(* IEC 61131-3 sources: Elmo_Master/Lasal_PRG/Welcon8Axis_EtherCAT_Test_With_RobotAxis/Network/HW_Network, 1 file *)

(* ---- ONE_HW_Network_Table.st ---- *)
#define OBJECTS_CONFIG

//Define part of class _SyncMeasure
#define _SYNCM_PLLLOCK_MASK 2#11110000
#define _SYNCM_PLLLOCK      2#10100000

#define _SYNCM_PLLLOCK_MASK_MASTER 2#11000000
#define _SYNCM_PLLLOCK_MASTER      2#10000000

#define _SYNCM_PLLLOCK_MASK_OWN 2#00110000
#define _SYNCM_PLLLOCK_OWN      2#00100000

#define _SYNCM_PLL_DELTAREG_ENABLE   2#01001000
#define _SYNCM_PLL_DELTAREG_DISABLE  2#01000000

#define _SYNCM_25US 2500 // [10 ns]
#define _SYNCM_50US 5000 // [10 ns]

// #define _SYNCM_DEBUG
#include "..\..\source\interfaces\lsl_st_pll.h"
#include "..\..\Source\BusInterface.h"
//Define part of class _SyncMeasureECAT
#define _SYNCMCAT_MAX_FILTER_SIZE 100

//#define _SYNCMECAT_DEBUG

#define _SYNCMECAT_FilterSize_LL_Measure_Delta   150
#define _SYNCMECAT_FilterSize_LLFP_Offset         25
#define _SYNCMECAT_FilterSize_LL_Roundtrip       500
#define _SYNCMECAT_FilterSize_RCLL_Offset         10
#define _SYNCMECAT_FilterSize_Deltatime           10
#define _SYNCMECAT_FilterSize_Gradient            30
#define _SYNCMECAT_FilterSize_Corr_Steig          80

#define _SYNCMECAT_DCSlvM_AdjustLevel             1//10 //ns

#define _SYNCMECAT_SyncStart_CorrFactorUp        100
#define _SYNCMECAT_SyncStart_CorrFactorDown       50

#define _SYNCMECAT_SyncStart_CorrFactorUp_fine     1
#define _SYNCMECAT_SyncStart_CorrFactorDown_fine   1

#define _SYNCMECAT_SyncStart_DistFactUp        25000
#define _SYNCMECAT_SyncStart_DistFactDown      25000
#include "..\..\Class\ECAT_Master_Base\ECAT_Master_Base.h"
#include "..\..\Class\_SyncMeasureECAT\_64BitTimestamp.h"
//Define part of class BusInterfaceSDIASInternal
#define BUSIF_INTERNAL_MAX_NR_DO 100

// Defines for Mutex Generation
#define INTERNAL_STR_MUTEX_NAME_SEPERATOR ".."
#define INTERNAL_MUTEX_NAME_END_LENGTH 5
#define INTERNAL_MUTEX_NAME_MAX_LENGTH 32
#include "..\..\Source\interfaces\lsl_st_mt.h"
#include "..\..\Class\HwControl\HwControl.h"
#include "..\..\Source\interfaces\lsl_st_hardwaretree.h"
//Define part of class ECAT_Slave_Base
#define ECAT_SB_SDO_LOCK                    16#A1B2C3D4
#define ECAT_SB_SDO_FREE                    16#E5F60718

#define ECAT_SB_VENDORID_SIGMATEK           16#000088FA

//CoE Communication area
#define ECAT_SB_INDEX_DEVICE_TYPE           16#1000 //mandatory
#define ECAT_SB_SUBINDEX_DEVICE_TYPE              0

#define ECAT_SB_INDEX_DEVICE_NAME           16#1008 //optional
#define ECAT_SB_SUBINDEX_DEVICE_NAME              0

#define ECAT_SB_INDEX_HARDWARE_VERSION      16#1009 //optional
#define ECAT_SB_SUBINDEX_HARDWARE_VERSION         0

#define ECAT_SB_INDEX_SOFTWARE_VERSION      16#100A //optional
#define ECAT_SB_SUBINDEX_SOFTWARE_VERSION         0

#define ECAT_SB_INDEX_IDENTITY_OBJECT       16#1018 //mandatory
#define ECAT_SB_SUBINDEX_IDENTITY_OBJECT          0

#define ECAT_SB_DEFAULT_SDO_TIMEOUT         2000

#define ECAT_SB_PHYSICAL_START_ADRESS        1001
#include "..\..\Class\ECAT_Slave_Base\ECAT_Slave_Base.h"
#include "..\..\Source\interfaces\lsl_st_ecatm.h"
//Define part of class ECAT_DS402Base
// As defined in ETG.6010 D (R) V1.1.0

// PDO idx
#define ECAT_DS402BASE_IDX_CONTROLWORD  0x6040
#define ECAT_DS402BASE_IDX_STATUSWORD   0x6041

#define ECAT_DS402BASE_IDX_SETSPEED     0x60FF
#define ECAT_DS402BASE_IDX_ACTSPEED     0x606C

#define ECAT_DS402BASE_IDX_SETPOS       0x607A
#define ECAT_DS402BASE_IDX_ACTPOS       0x6064

#define ECAT_DS402BASE_IDX_ACTTORQUE    0x6077
#define ECAT_DS402BASE_IDX_SETTORQUE    0x6071

#define ECAT_DS402BASE_IDX_ACTXW        0x60F4
#include "..\..\Source\DriveSafetyIF.h"
//Define part of class ECAT_Master_Base
#define ECATM_MAX_NO_TASKS 5
#define ECATM_INC_CYC_CALLBACKS 5

#define ECATM_STR_ENI_FILE    "C:/lslsys/hwoutput.conf"      //Standard path of ENI-File

#define ECATM_MAX_VALUE_MISSING_FRAME_BEHAVIOUR 31
#define ECATM_MAX_SIZE_FRAME_ERROR_LOGBUFFER    50

#define ECATM_THREAD_PRIO_DISABLE               10 // Background
#define ECATM_THREAD_STACKSIZE              0x4000
#include "..\..\Source\interfaces\lsl_st_systrace.h"
#include "..\..\Source\interfaces\lsl_st_gpio.h"
#include "..\..\Source\interfaces\lsl_st_mediaplayer.h"
#include "..\..\Source\interfaces\lsl_st_pci.h"
#include "..\..\Source\interfaces\lsl_st_powermanagement.h"
#include "..\..\Source\interfaces\lsl_st_pwm.h"
#include "..\..\source\interfaces\lsl_st_spi.h"
#include "..\..\Source\interfaces\lsl_st_sysinfo.h"
#include "..\..\Source\interfaces\lsl_st_x_ram.h"
#include "..\..\Class\HwControl\watchdog.h"
#include "..\..\Class\HwControl\_HWKScope.h"
#include "..\..\Class\HwControl\HwControlParameters.h"
#include <.\lsl_st_mt.h>
//Define part of class SafetyUDP
#define SAFETY_UDP_MAX_SOCKETS                6     // Max number of socket

#define SAFETY_UDP_CLT_SEND_OK                0    // Send ok
#define SAFETY_UDP_CLT_INVALID_HANDLE        -1    // Invalid handle
#define SAFETY_UDP_CLT_NOT_OPEN              -2    // Socket is not open
#define SAFETY_UDP_CLT_SEND_FAILED           -3    // Send failed
#define SAFETY_UDP_CLT_SEND_BUFFER_FULL      -4    // Send buffer is full
#define SAFETY_UDP_CLT_DATA_TO_BIG           -5    // Data to big

#define SAFETY_UDP_MAXIMUM_SEGMENT_SIZE    1452    // Maximum of user data

#define SAFETY_UDP_TIMEOUT_OPENSOCKET    (1000)    //timeout for opening socket

#define SAFETY_UDP_RECEIVE_TIMEOUT          800

#define SAFETY_UDP_TX_BUFFER_SIZE          1024
//Define part of class SafetyManager
#define SM_LogBufferSize 1000
#define SM_MaxObjNameLen  256
#include "..\..\Class\SafetyManager\SafetyManager.h"
#include "..\..\Source\interfaces\lsl_st_safetydll.h"
//Define part of class SafetyRoutingTables
#define SRT_MAXIDX 15 // Currently there are 2 Tables for each Eni File / EtherMaster
//Define part of class SdiasManager
#define SDIAS_SDO_MAX_LENGTH              128
#define SDIAS_SDO_RINGBUFFER_NO            64
#define SDIAS_SDO_CHANNEL_NO                3   // fixed in the VI hardware to be 3

// watchdog trigger interval (after 130ms of no trigger the SDIAS HW goes into reset again and takes at least another 10ms to be ready again)
#define SDIAS_WATCHDOG_TRIGGER_TIME        40

// time needed by sdias modules to start up after the watchdog is triggered the first time in ms
#define SDIAS_HARDWARE_STARTUP_TIME        15

// sdias manager needs 2 ticks to handle event for read task (measure sync time)
#define SDIAS_SYNC_MEASURE_TICKS            2

// after activating the PLL SyncOut it takes 3 cycles until the SDIAS sync can be injected
#define SDIAS_CYCLES_WAIT_AFTER_SYNC_ENABLE 3

// wait 1 bus cycle at start to get valid numbers in the task info
#define SDIAS_TASKINFO_READY_TICKS          1

// time to wait (in ms) until other tasks in the same or lower priority than post init have done their stuff
#define SDIAS_WAIT_TIME_IN_POST_INIT        1

#define SIZE_PER_SDIAS_CLIENT               16#0400

// for far memory accesses: 1 module can hold maximum 256 1K blocks (0-255)
#define SDIAS_1K_BLOCK_NO                       256

// far memory accesses maximum length in bytes
#define SDIAS_MAX_SIZE_FAR_MEM_ACCESS           127

#define SDIAS_OFFSET_HW_CONFIG              16#FF00
#define SDIAS_OFFSET_TASK_EVENT_IDS         16#FF10
#define SDIAS_OFFSET_FEATURE_INFO           16#FF18
#define SDIAS_OFFSET_APPLI_LED_STATES       16#FF20
#define SDIAS_OFFSET_SYNC_INJECTION_CFG     16#FF3D
#define SDIAS_OFFSET_TRIGGER_UNIT_SETUP_0   16#FF41
#define SDIAS_OFFSET_TRIGGER_UNIT_SETUP_1   16#FF45
#define SDIAS_OFFSET_TASK_START_CFG_0       16#FF60
#define SDIAS_OFFSET_TASK_CONFIG_0          16#FF86
#define SDIAS_OFFSET_TASK_CONFIG_1          16#FF96
#define SDIAS_OFFSET_TASK_INFO_1            16#FF94
#define SDIAS_OFFSET_TASK_HANDSHAKE_1       16#FF9B
#define SDIAS_OFFSET_TASK_DURATION_TIME_1   16#FF9C
#define SDIAS_OFFSET_TASK_DURATION_TIME_2   16#FFAC
#define SDIAS_OFFSET_TASK_CONFIG_2          16#FFA6

#define SDIAS_RETRIES_ALLOWED         2

// mask to get global error flag out of message counter byte of SDO responses
#define SDIAS_MASK_GLOBAL_ERROR_FLAG        16#80

// mask to get message counter out of message counter byte of SDO responses
#define SDIAS_MASK_MESSAGE_COUNTER          16#3F

#define SDIAS_EVENT_MASK_ID_SYNC_OUT0       16#10
#define SDIAS_EVENT_MASK_ID_SYNC_OUT1       16#11
#define SDIAS_EVENT_MASK_ID_SYNC_OUT2       16#12
#define SDIAS_EVENT_MASK_ID_SYNC_OUT3       16#13

#define SDIAS_MANAGER_SYNC_SYNCOUT_ID       16#85
#define SDIAS_TASK_START_EVENT_SYNCOUT_ID   16#86

#define SDIAS_PLACE_NO_MODULE_ADDED_SO_FAR  16#80000000

#define SDIAS_TRIGGER_UNIT_BYTE_SIZE        2

#define SDIAS_WAIT_TIME_FIRMWARE_HANDSHAKE  5 * 1000

// if the firmware version is below this, there might be problems with SCP111 and other modules => print warning at startup
#define SDIAS_FW_VERSION_SDO_ERROR_FIXED    16#120

// if the protocol version ist below this, Control Read/Broadcast Write Command is not supported by sdiasmanager
#define SDIAS_PROTOCOLVERSION_BROADCAST     16#120

// if the cil version ist below this, Control Read/Broadcast Write Command is not supported by OS for local SDIAS.
#define SDIAS_CILVERSION_BROADCAST         16#5001

// timeout for blocking the init during initialisation (in ms)
#define SDIAS_INIT_BLOCK_TIMEOUT            20 * 1000

#define SDIAS_MUTEX_NAME_END_LENGTH 3
#define SDIAS_MUTEX_NAME_MAX_LENGTH 32
#define SDIAS_MUTEX_STR_SEPERATOR   ".."

//#define SDIAS_RT_TIME_MEASUREMENT
#ifdef SDIAS_RT_TIME_MEASUREMENT
  #pragma message("ATTENTION: SDIAS real time measurement is active and needs additional ressources in the realtime task")
#endif

(* SDIAS data object commands  *)
#define	 SDIAS_CMD_END							  0x00			(* End command										          *)
#define	 SDIAS_CMD_ACC_MEMORY				  0x01			(* Access dpram memory								      *)
#define	 SDIAS_CMD_ACC_CONTROL				0x02			(* Access dpram control memory						  *)
#define	 SDIAS_CMD_GLOBAL						  0x03			(* SDIAS global command								      *)
#define	 SDIAS_CMD_COPY_LOCAL					0x04			(* DPRAM copy command in local dpram				*)
#define	 SDIAS_CMD_JMP_LOCAL					0x05			(* DPRAM jump command in local dpram 				*)
#define  SDIAS_CMD_ACC_MEMORY_FAR     0x07      (* SDIAS Far Memory Access                  *)

(* SDIAS defines for data object handling *)
// Write data oject list
#define	 SDIAS_DOL_WRITE_USAGE_DOL_EMPTY	  0x20			(* Usage of empty write dol list (wachtdog trigger + end command)   *)
#define	 SDIAS_DOL_WRITE_USAGE_DTA_EMPTY	  0x03			(* Usage of empty write dol data (DO ctrl of 2x copy command for task information + DO ctrl of watchdog trigger      *)
#define	 SDIAS_DOL_WRITE_OFFSET_END_CMD			0x10			(* One data object in list - offset = 1 DO size = 0x10						  *)
#define	 SDIAS_DOL_WRITE_OFFSET_FIRST_DTA		0x02			(* Offset of first data byte of second copy command = 2 (DO ctrl)   *)
#define	 SDIAS_DOL_WRITE_OFFSET_LAST_DTA		0x02			(* Offset of last data byte of second copy command = 2 (DO ctrl )   *)

// Read data oject list
#define	 SDIAS_DOL_READ_USAGE_DOL_EMPTY	    0x30			(* Usage of empty read dol list (2x task info copy command + end command)   *)
#define	 SDIAS_DOL_READ_USAGE_DTA_EMPTY	    0x0D			(* Usage of empty write dol data (DO ctrl of 2x copy command for task information + DO ctrl of watchdog trigger      *)
#define	 SDIAS_DOL_READ_OFFSET_END_CMD			0x20			(* One data object in list - offset = 1 DO size = 0x10						          *)
#define	 SDIAS_DOL_READ_OFFSET_FIRST_DTA		0x07			(* Offset of first data byte of second copy command = 7 = DO state          *)
#define	 SDIAS_DOL_READ_OFFSET_LAST_DTA		  0x0C			(* Offset of last data byte of second copy command = 12 (last byte of task information)       *)

//Versionsnumber where SDIAS SPI Read Accesses are available
#define  SDIAS_SDO_SPI_FIRMWARE_VERSION_AVAILABLE 16#0120

//error info mask
#define  SDIAS_ERROR_INFO_MASK    2#1000011000011111

// Broadcast DO Info
#define SDIAS_OFFSET_CLIENT_CTRLTIMESTAMP   16#0190
#define SDIAS_NR_TIMEBROADCAST_DOS 2
#define SDIAS_TIMEBROADCAST_SUBCMD 16#B0
#include "..\..\Class\SdiasManager\SdiasManager.h"
//Define part of class SdiasPLC
#define SDIASM_OBJECT_PATH            16#88000002   // Object Path for VSDIASmanager Length = 2 (First 2byte), Domain = 0 (3rd byte), Escape Sequence SDIAS (4th byte)
//Define part of class VaranManager
#define SIZE_PAYLOAD_FRAME_HEADER_DO      16#38  // Const because datasize is in the Payload DOs
#define SIZE_PAYLOAD_IRQ_FRAME_HEADER_DO  16#40  // Const because datasize is in the Payload DOs

#define VM_MAX_POST_INIT_MODULES  1000

#define VM_OBJECT_PATH            16#81000002   // Object Path for Varanmanager Length = 2 (First 2byte), Domain = 0 (3rd byte), Escape Sequence Varan (4th byte)
#include "..\..\Class\VaranManager\VaranManager.h"
#include "..\..\Source\interfaces\lsl_st_kernel.h"
//Define part of class WELCON_1
//{{ECAT_DEFINES
#define WELCON_1_ETHERCATSLAVE_PRODUCT_CODE 536870913
#define WELCON_1_ETHERCATSLAVE_VENDOR_ID    2985
#define WELCON_1_CONTROLWORD_INDEX		16#6040
#define WELCON_1_CONTROLWORD_SUBINDEX			0
#define WELCON_1_SETPOS_INDEX		16#607A
#define WELCON_1_SETPOS_SUBINDEX			0
#define WELCON_1_SETSPEED_INDEX		16#60FF
#define WELCON_1_SETSPEED_SUBINDEX			0
#define WELCON_1_SETTORQUE_INDEX		16#6071
#define WELCON_1_SETTORQUE_SUBINDEX			0
#define WELCON_1_RXPDO9_PHYSICALOUTPUTS1_INDEX		16#60FE
#define WELCON_1_RXPDO9_PHYSICALOUTPUTS1_SUBINDEX			1
#define WELCON_1_RXPDO9_MODESOFOPERATION1_INDEX		16#6060
#define WELCON_1_RXPDO9_MODESOFOPERATION1_SUBINDEX			0
#define WELCON_1_RXPDO9_CONTROLWORD2_INDEX		16#6840
#define WELCON_1_RXPDO9_CONTROLWORD2_SUBINDEX			0
#define WELCON_1_RXPDO9_TARGETPOSITION2_INDEX		16#687A
#define WELCON_1_RXPDO9_TARGETPOSITION2_SUBINDEX			0
#define WELCON_1_RXPDO9_TARGETVELOCITY2_INDEX		16#68FF
#define WELCON_1_RXPDO9_TARGETVELOCITY2_SUBINDEX			0
#define WELCON_1_RXPDO9_TARGETTORQUE2_INDEX		16#6871
#define WELCON_1_RXPDO9_TARGETTORQUE2_SUBINDEX			0
#define WELCON_1_RXPDO9_PHYSICALOUTPUTS2_INDEX		16#68FE
#define WELCON_1_RXPDO9_PHYSICALOUTPUTS2_SUBINDEX			1
#define WELCON_1_RXPDO9_MODESOFOPERATION2_INDEX		16#6860
#define WELCON_1_RXPDO9_MODESOFOPERATION2_SUBINDEX			0
#define WELCON_1_STATEWORD_INDEX		16#6041
#define WELCON_1_STATEWORD_SUBINDEX			0
#define WELCON_1_ACTPOS_INDEX		16#6064
#define WELCON_1_ACTPOS_SUBINDEX			0
#define WELCON_1_ACTSPEED_INDEX		16#606C
#define WELCON_1_ACTSPEED_SUBINDEX			0
#define WELCON_1_ACTTORQUE_INDEX		16#6077
#define WELCON_1_ACTTORQUE_SUBINDEX			0
#define WELCON_1_TXPDO9_DIGITALINPUTS1_INDEX		16#60FD
#define WELCON_1_TXPDO9_DIGITALINPUTS1_SUBINDEX			0
#define WELCON_1_TXPDO9_MODESOFOPERATIONDISPLAY1_INDEX		16#6061
#define WELCON_1_TXPDO9_MODESOFOPERATIONDISPLAY1_SUBINDEX			0
#define WELCON_1_TXPDO9_STATUSWORD2_INDEX		16#6841
#define WELCON_1_TXPDO9_STATUSWORD2_SUBINDEX			0
#define WELCON_1_TXPDO9_POSITIONACTUALVALUE2_INDEX		16#6864
#define WELCON_1_TXPDO9_POSITIONACTUALVALUE2_SUBINDEX			0
#define WELCON_1_TXPDO9_VELOCITYACTUALVALUE2_INDEX		16#686C
#define WELCON_1_TXPDO9_VELOCITYACTUALVALUE2_SUBINDEX			0
#define WELCON_1_TXPDO9_TORQUEACTUALVALUE2_INDEX		16#6877
#define WELCON_1_TXPDO9_TORQUEACTUALVALUE2_SUBINDEX			0
#define WELCON_1_TXPDO9_DIGITALINPUTS2_INDEX		16#68FD
#define WELCON_1_TXPDO9_DIGITALINPUTS2_SUBINDEX			0
#define WELCON_1_TXPDO9_MODESOFOPERATIONDISPLAY2_INDEX		16#6861
#define WELCON_1_TXPDO9_MODESOFOPERATIONDISPLAY2_SUBINDEX			0
//}}ECAT_DEFINES
//Define part of class WELCON_2
//{{ECAT_DEFINES
#define WELCON_2_ETHERCATSLAVE_PRODUCT_CODE 536870913
#define WELCON_2_ETHERCATSLAVE_VENDOR_ID    2985
#define WELCON_2_CONTROLWORD_INDEX		16#6040
#define WELCON_2_CONTROLWORD_SUBINDEX			0
#define WELCON_2_SETPOS_INDEX		16#607A
#define WELCON_2_SETPOS_SUBINDEX			0
#define WELCON_2_SETSPEED_INDEX		16#60FF
#define WELCON_2_SETSPEED_SUBINDEX			0
#define WELCON_2_SETTORQUE_INDEX		16#6071
#define WELCON_2_SETTORQUE_SUBINDEX			0
#define WELCON_2_RXPDO9_PHYSICALOUTPUTS1_INDEX		16#60FE
#define WELCON_2_RXPDO9_PHYSICALOUTPUTS1_SUBINDEX			1
#define WELCON_2_RXPDO9_MODESOFOPERATION1_INDEX		16#6060
#define WELCON_2_RXPDO9_MODESOFOPERATION1_SUBINDEX			0
#define WELCON_2_RXPDO9_CONTROLWORD2_INDEX		16#6840
#define WELCON_2_RXPDO9_CONTROLWORD2_SUBINDEX			0
#define WELCON_2_RXPDO9_TARGETPOSITION2_INDEX		16#687A
#define WELCON_2_RXPDO9_TARGETPOSITION2_SUBINDEX			0
#define WELCON_2_RXPDO9_TARGETVELOCITY2_INDEX		16#68FF
#define WELCON_2_RXPDO9_TARGETVELOCITY2_SUBINDEX			0
#define WELCON_2_RXPDO9_TARGETTORQUE2_INDEX		16#6871
#define WELCON_2_RXPDO9_TARGETTORQUE2_SUBINDEX			0
#define WELCON_2_RXPDO9_PHYSICALOUTPUTS2_INDEX		16#68FE
#define WELCON_2_RXPDO9_PHYSICALOUTPUTS2_SUBINDEX			1
#define WELCON_2_RXPDO9_MODESOFOPERATION2_INDEX		16#6860
#define WELCON_2_RXPDO9_MODESOFOPERATION2_SUBINDEX			0
#define WELCON_2_STATEWORD_INDEX		16#6041
#define WELCON_2_STATEWORD_SUBINDEX			0
#define WELCON_2_ACTPOS_INDEX		16#6064
#define WELCON_2_ACTPOS_SUBINDEX			0
#define WELCON_2_ACTSPEED_INDEX		16#606C
#define WELCON_2_ACTSPEED_SUBINDEX			0
#define WELCON_2_ACTTORQUE_INDEX		16#6077
#define WELCON_2_ACTTORQUE_SUBINDEX			0
#define WELCON_2_TXPDO9_DIGITALINPUTS1_INDEX		16#60FD
#define WELCON_2_TXPDO9_DIGITALINPUTS1_SUBINDEX			0
#define WELCON_2_TXPDO9_MODESOFOPERATIONDISPLAY1_INDEX		16#6061
#define WELCON_2_TXPDO9_MODESOFOPERATIONDISPLAY1_SUBINDEX			0
#define WELCON_2_TXPDO9_STATUSWORD2_INDEX		16#6841
#define WELCON_2_TXPDO9_STATUSWORD2_SUBINDEX			0
#define WELCON_2_TXPDO9_POSITIONACTUALVALUE2_INDEX		16#6864
#define WELCON_2_TXPDO9_POSITIONACTUALVALUE2_SUBINDEX			0
#define WELCON_2_TXPDO9_VELOCITYACTUALVALUE2_INDEX		16#686C
#define WELCON_2_TXPDO9_VELOCITYACTUALVALUE2_SUBINDEX			0
#define WELCON_2_TXPDO9_TORQUEACTUALVALUE2_INDEX		16#6877
#define WELCON_2_TXPDO9_TORQUEACTUALVALUE2_SUBINDEX			0
#define WELCON_2_TXPDO9_DIGITALINPUTS2_INDEX		16#68FD
#define WELCON_2_TXPDO9_DIGITALINPUTS2_SUBINDEX			0
#define WELCON_2_TXPDO9_MODESOFOPERATIONDISPLAY2_INDEX		16#6861
#define WELCON_2_TXPDO9_MODESOFOPERATIONDISPLAY2_SUBINDEX			0
//}}ECAT_DEFINES
//Define part of class WELCON_3
//{{ECAT_DEFINES
#define WELCON_3_ETHERCATSLAVE_PRODUCT_CODE 536870913
#define WELCON_3_ETHERCATSLAVE_VENDOR_ID    2985
#define WELCON_3_CONTROLWORD_INDEX		16#6040
#define WELCON_3_CONTROLWORD_SUBINDEX			0
#define WELCON_3_SETPOS_INDEX		16#607A
#define WELCON_3_SETPOS_SUBINDEX			0
#define WELCON_3_SETSPEED_INDEX		16#60FF
#define WELCON_3_SETSPEED_SUBINDEX			0
#define WELCON_3_SETTORQUE_INDEX		16#6071
#define WELCON_3_SETTORQUE_SUBINDEX			0
#define WELCON_3_RXPDO9_PHYSICALOUTPUTS1_INDEX		16#60FE
#define WELCON_3_RXPDO9_PHYSICALOUTPUTS1_SUBINDEX			1
#define WELCON_3_RXPDO9_MODESOFOPERATION1_INDEX		16#6060
#define WELCON_3_RXPDO9_MODESOFOPERATION1_SUBINDEX			0
#define WELCON_3_RXPDO9_CONTROLWORD2_INDEX		16#6840
#define WELCON_3_RXPDO9_CONTROLWORD2_SUBINDEX			0
#define WELCON_3_RXPDO9_TARGETPOSITION2_INDEX		16#687A
#define WELCON_3_RXPDO9_TARGETPOSITION2_SUBINDEX			0
#define WELCON_3_RXPDO9_TARGETVELOCITY2_INDEX		16#68FF
#define WELCON_3_RXPDO9_TARGETVELOCITY2_SUBINDEX			0
#define WELCON_3_RXPDO9_TARGETTORQUE2_INDEX		16#6871
#define WELCON_3_RXPDO9_TARGETTORQUE2_SUBINDEX			0
#define WELCON_3_RXPDO9_PHYSICALOUTPUTS2_INDEX		16#68FE
#define WELCON_3_RXPDO9_PHYSICALOUTPUTS2_SUBINDEX			1
#define WELCON_3_RXPDO9_MODESOFOPERATION2_INDEX		16#6860
#define WELCON_3_RXPDO9_MODESOFOPERATION2_SUBINDEX			0
#define WELCON_3_STATEWORD_INDEX		16#6041
#define WELCON_3_STATEWORD_SUBINDEX			0
#define WELCON_3_ACTPOS_INDEX		16#6064
#define WELCON_3_ACTPOS_SUBINDEX			0
#define WELCON_3_ACTSPEED_INDEX		16#606C
#define WELCON_3_ACTSPEED_SUBINDEX			0
#define WELCON_3_ACTTORQUE_INDEX		16#6077
#define WELCON_3_ACTTORQUE_SUBINDEX			0
#define WELCON_3_TXPDO9_DIGITALINPUTS1_INDEX		16#60FD
#define WELCON_3_TXPDO9_DIGITALINPUTS1_SUBINDEX			0
#define WELCON_3_TXPDO9_MODESOFOPERATIONDISPLAY1_INDEX		16#6061
#define WELCON_3_TXPDO9_MODESOFOPERATIONDISPLAY1_SUBINDEX			0
#define WELCON_3_TXPDO9_STATUSWORD2_INDEX		16#6841
#define WELCON_3_TXPDO9_STATUSWORD2_SUBINDEX			0
#define WELCON_3_TXPDO9_POSITIONACTUALVALUE2_INDEX		16#6864
#define WELCON_3_TXPDO9_POSITIONACTUALVALUE2_SUBINDEX			0
#define WELCON_3_TXPDO9_VELOCITYACTUALVALUE2_INDEX		16#686C
#define WELCON_3_TXPDO9_VELOCITYACTUALVALUE2_SUBINDEX			0
#define WELCON_3_TXPDO9_TORQUEACTUALVALUE2_INDEX		16#6877
#define WELCON_3_TXPDO9_TORQUEACTUALVALUE2_SUBINDEX			0
#define WELCON_3_TXPDO9_DIGITALINPUTS2_INDEX		16#68FD
#define WELCON_3_TXPDO9_DIGITALINPUTS2_SUBINDEX			0
#define WELCON_3_TXPDO9_MODESOFOPERATIONDISPLAY2_INDEX		16#6861
#define WELCON_3_TXPDO9_MODESOFOPERATIONDISPLAY2_SUBINDEX			0
//}}ECAT_DEFINES
//Define part of class WELCON_4
//{{ECAT_DEFINES
#define WELCON_4_ETHERCATSLAVE_PRODUCT_CODE 536870913
#define WELCON_4_ETHERCATSLAVE_VENDOR_ID    2985
#define WELCON_4_CONTROLWORD_INDEX		16#6040
#define WELCON_4_CONTROLWORD_SUBINDEX			0
#define WELCON_4_SETPOS_INDEX		16#607A
#define WELCON_4_SETPOS_SUBINDEX			0
#define WELCON_4_SETSPEED_INDEX		16#60FF
#define WELCON_4_SETSPEED_SUBINDEX			0
#define WELCON_4_SETTORQUE_INDEX		16#6071
#define WELCON_4_SETTORQUE_SUBINDEX			0
#define WELCON_4_RXPDO9_PHYSICALOUTPUTS1_INDEX		16#60FE
#define WELCON_4_RXPDO9_PHYSICALOUTPUTS1_SUBINDEX			1
#define WELCON_4_RXPDO9_MODESOFOPERATION1_INDEX		16#6060
#define WELCON_4_RXPDO9_MODESOFOPERATION1_SUBINDEX			0
#define WELCON_4_RXPDO9_CONTROLWORD2_INDEX		16#6840
#define WELCON_4_RXPDO9_CONTROLWORD2_SUBINDEX			0
#define WELCON_4_RXPDO9_TARGETPOSITION2_INDEX		16#687A
#define WELCON_4_RXPDO9_TARGETPOSITION2_SUBINDEX			0
#define WELCON_4_RXPDO9_TARGETVELOCITY2_INDEX		16#68FF
#define WELCON_4_RXPDO9_TARGETVELOCITY2_SUBINDEX			0
#define WELCON_4_RXPDO9_TARGETTORQUE2_INDEX		16#6871
#define WELCON_4_RXPDO9_TARGETTORQUE2_SUBINDEX			0
#define WELCON_4_RXPDO9_PHYSICALOUTPUTS2_INDEX		16#68FE
#define WELCON_4_RXPDO9_PHYSICALOUTPUTS2_SUBINDEX			1
#define WELCON_4_RXPDO9_MODESOFOPERATION2_INDEX		16#6860
#define WELCON_4_RXPDO9_MODESOFOPERATION2_SUBINDEX			0
#define WELCON_4_STATEWORD_INDEX		16#6041
#define WELCON_4_STATEWORD_SUBINDEX			0
#define WELCON_4_ACTPOS_INDEX		16#6064
#define WELCON_4_ACTPOS_SUBINDEX			0
#define WELCON_4_ACTSPEED_INDEX		16#606C
#define WELCON_4_ACTSPEED_SUBINDEX			0
#define WELCON_4_ACTTORQUE_INDEX		16#6077
#define WELCON_4_ACTTORQUE_SUBINDEX			0
#define WELCON_4_TXPDO9_DIGITALINPUTS1_INDEX		16#60FD
#define WELCON_4_TXPDO9_DIGITALINPUTS1_SUBINDEX			0
#define WELCON_4_TXPDO9_MODESOFOPERATIONDISPLAY1_INDEX		16#6061
#define WELCON_4_TXPDO9_MODESOFOPERATIONDISPLAY1_SUBINDEX			0
#define WELCON_4_TXPDO9_STATUSWORD2_INDEX		16#6841
#define WELCON_4_TXPDO9_STATUSWORD2_SUBINDEX			0
#define WELCON_4_TXPDO9_POSITIONACTUALVALUE2_INDEX		16#6864
#define WELCON_4_TXPDO9_POSITIONACTUALVALUE2_SUBINDEX			0
#define WELCON_4_TXPDO9_VELOCITYACTUALVALUE2_INDEX		16#686C
#define WELCON_4_TXPDO9_VELOCITYACTUALVALUE2_SUBINDEX			0
#define WELCON_4_TXPDO9_TORQUEACTUALVALUE2_INDEX		16#6877
#define WELCON_4_TXPDO9_TORQUEACTUALVALUE2_SUBINDEX			0
#define WELCON_4_TXPDO9_DIGITALINPUTS2_INDEX		16#68FD
#define WELCON_4_TXPDO9_DIGITALINPUTS2_SUBINDEX			0
#define WELCON_4_TXPDO9_MODESOFOPERATIONDISPLAY2_INDEX		16#6861
#define WELCON_4_TXPDO9_MODESOFOPERATIONDISPLAY2_SUBINDEX			0
//}}ECAT_DEFINES

FUNCTION GLOBAL TAB ONE_HW_Network
-1$UINT, 0$UINT,
0$UINT, 0$UINT,

38$UDINT,
TO_UDINT(529317953), "_CanLib", 1$UINT, 11$UINT, 2$UINT,
TO_UDINT(4078275645), "_SerLib", 1$UINT, 36$UINT, 3$UINT,
TO_UDINT(34287727), "_SyncMeasure", 1$UINT, 4$UINT, 0$UINT,
TO_UDINT(820122881), "_SyncMeasureECAT", 1$UINT, 3$UINT, 1$UINT,
TO_UDINT(2897291062), "ASCII_BIN", 1$UINT, 21$UINT, 1$UINT,
TO_UDINT(3882880897), "BusInterfaceSDIASInternal", 2$UINT, 2$UINT, 0$UINT,
TO_UDINT(2377812740), "CP313_IOs", 1$UINT, 1$UINT, 1$UINT,
TO_UDINT(794617671), "CriticalSection", 0$UINT, 4$UINT, 2$UINT,
TO_UDINT(861770287), "ECAT_DS402Base", 1$UINT, 2$UINT, 0$UINT,
TO_UDINT(4097056936), "ECAT_Master_Base", 2$UINT, 3$UINT, 0$UINT,
TO_UDINT(1515440174), "ECAT_Slave_Base", 2$UINT, 1$UINT, 0$UINT,
TO_UDINT(1021147964), "EtherCAT_Hub_Base", 1$UINT, 2$UINT, 5$UINT,
TO_UDINT(631677903), "EtherCAT_PLC", 2$UINT, 2$UINT, 1$UINT,
TO_UDINT(1916923939), "GetCILInterface", 1$UINT, 5$UINT, 6$UINT,
TO_UDINT(3238133653), "Hub_Base", 1$UINT, 22$UINT, 0$UINT,
TO_UDINT(1770276445), "Hub_Base_Root", 2$UINT, 12$UINT, 1$UINT,
TO_UDINT(3078259981), "HwcLogging", 1$UINT, 1$UINT, 1$UINT,
TO_UDINT(2471641665), "HwControl", 6$UINT, 0$UINT, 1$UINT,
TO_UDINT(1193052171), "HwControlBase", 1$UINT, 11$UINT, 0$UINT,
TO_UDINT(4260294091), "HWRtPostScan", 1$UINT, 1$UINT, 1$UINT,
TO_UDINT(2225119864), "MerkerEx", 1$UINT, 22$UINT, 9$UINT,
TO_UDINT(1799751072), "SafetyManager", 3$UINT, 0$UINT, 1$UINT,
TO_UDINT(3387336038), "SafetyRoutingTables", 1$UINT, 0$UINT, 1$UINT,
TO_UDINT(3727715967), "SafetyUDP", 1$UINT, 5$UINT, 0$UINT,
TO_UDINT(4173303375), "SdiasHubBase", 1$UINT, 11$UINT, 1$UINT,
TO_UDINT(2118381352), "SdiasManager", 1$UINT, 100$UINT, 1$UINT,
TO_UDINT(1159122596), "SdiasPLC", 2$UINT, 8$UINT, 1$UINT,
TO_UDINT(1850111279), "String", 1$UINT, 11$UINT, 9$UINT,
TO_UDINT(2898603620), "StringInternal", 1$UINT, 86$UINT, 0$UINT,
TO_UDINT(2940693151), "VaranManager", 3$UINT, 9$UINT, 0$UINT,
TO_UDINT(1989862026), "VaranManager_1", 2$UINT, 8$UINT, 1$UINT,
TO_UDINT(4035182347), "VaranManager_Base", 1$UINT, 27$UINT, 0$UINT,
TO_UDINT(3232495061), "VirtualBaseInit", 1$UINT, 3$UINT, 0$UINT,
TO_UDINT(2662678246), "WELCON_1", 0$UINT, 0$UINT, 1$UINT,
TO_UDINT(129789788), "WELCON_2", 0$UINT, 0$UINT, 1$UINT,
TO_UDINT(1891327946), "WELCON_3", 0$UINT, 0$UINT, 1$UINT,
TO_UDINT(4007643753), "WELCON_4", 0$UINT, 0$UINT, 1$UINT,
TO_UDINT(819479645), "XXXBase_IOs", 1$UINT, 4$UINT, 0$UINT,

1$UINT, TO_UDINT(3425326136), "CP313_IOS1\_BASE\_CANLIB1",
1$UINT, TO_UDINT(1428358530), "CP313_IOS1\_BASE\_CANLIB2",

1$UINT, TO_UDINT(2507534435), "CP313_IOS1\_BASE\_SERLIB1",
1$UINT, TO_UDINT(209494489), "CP313_IOS1\_BASE\_SERLIB2",
1$UINT, TO_UDINT(2071695695), "CP313_IOS1\_BASE\_SERLIB3",

1$UINT, TO_UDINT(1058685178), "ETHERCAT_PLC1\_BASE\_SYNCMEASUREECAT1",

1$UINT, TO_UDINT(3603645853), "VARANMANAGER_11\_BASE\ASCII_BIN1",

_NO_ATTR, TO_UDINT(2218561829), "CP313_IOS1",

1$UINT, TO_UDINT(2972590922), "HWCONTROL1\SAFETYMANAGER\UDPRECEIVEDATA",
1$UINT, TO_UDINT(1868223583), "HWCONTROL1\SAFETYMANAGER\UDPSENDDATA",

1$UINT, TO_UDINT(4288059666), "ETHERCAT_PLC1\ETHERCAT_HUB_BASE1",
1$UINT, TO_UDINT(187678911), "WELCON_11\ETHERCAT_HUB_BASE_1",
1$UINT, TO_UDINT(844590591), "WELCON_21\ETHERCAT_HUB_BASE_1",
1$UINT, TO_UDINT(629082431), "WELCON_31\ETHERCAT_HUB_BASE_1",
1$UINT, TO_UDINT(1084635007), "WELCON_41\ETHERCAT_HUB_BASE_1",

_NO_ATTR, TO_UDINT(2283968053), "ETHERCAT_PLC1",

1$UINT, TO_UDINT(2153717368), "ETHERCAT_PLC1\_BASE\GETCILINTERFACE_ECAT",
1$UINT, TO_UDINT(3141338546), "ETHERCAT_PLC1\_BASE\_SYNCMEASUREECAT1\_BASE\GETCILINTERFACEPLL",
1$UINT, TO_UDINT(4138461647), "WELCON_11\_BASE\_BASE\GETCILINTERFACE_ECAT",
1$UINT, TO_UDINT(2105071574), "WELCON_21\_BASE\_BASE\GETCILINTERFACE_ECAT",
1$UINT, TO_UDINT(3001466910), "WELCON_31\_BASE\_BASE\GETCILINTERFACE_ECAT",
1$UINT, TO_UDINT(2981080485), "WELCON_41\_BASE\_BASE\GETCILINTERFACE_ECAT",

1$UINT, TO_UDINT(1776428101), "VARANMANAGER_11\HUB_BASE_ROOT0",

1$UINT, TO_UDINT(3105254819), "HWCONTROL1\HWCLOGGING",

_NO_ATTR, TO_UDINT(2190789875), "HWCONTROL1",

1$UINT, TO_UDINT(1673205898), "HWCONTROL1\HWRTPOSTSCAN",

1$UINT, TO_UDINT(2768321018), "ETHERCAT_PLC1\_BASE\STRSOFTWAREVERSION\MERKEREX0",
1$UINT, TO_UDINT(1103896242), "WELCON_11\_BASE\_BASE\DEVICENAMESTR\MERKEREX0",
1$UINT, TO_UDINT(1954235937), "WELCON_11\_BASE\_BASE\PRODUCTREVSTR\MERKEREX0",
1$UINT, TO_UDINT(203693781), "WELCON_21\_BASE\_BASE\DEVICENAMESTR\MERKEREX0",
1$UINT, TO_UDINT(965953094), "WELCON_21\_BASE\_BASE\PRODUCTREVSTR\MERKEREX0",
1$UINT, TO_UDINT(2175591223), "WELCON_31\_BASE\_BASE\DEVICENAMESTR\MERKEREX0",
1$UINT, TO_UDINT(3021716388), "WELCON_31\_BASE\_BASE\PRODUCTREVSTR\MERKEREX0",
1$UINT, TO_UDINT(2549358107), "WELCON_41\_BASE\_BASE\DEVICENAMESTR\MERKEREX0",
1$UINT, TO_UDINT(2722317960), "WELCON_41\_BASE\_BASE\PRODUCTREVSTR\MERKEREX0",

1$UINT, TO_UDINT(1778590035), "HWCONTROL1\SAFETYMANAGER",

1$UINT, TO_UDINT(209976428), "HWCONTROL1\SAFETYMANAGER\SAFETYROUTINGTABLES1",

1$UINT, TO_UDINT(1007630054), "SDIASPLC1\SDIASHUBBASE1",

1$UINT, TO_UDINT(4015996540), "SDIASPLC1\SDIASMANAGER1",

_NO_ATTR, TO_UDINT(1378000520), "SDIASPLC1",

1$UINT, TO_UDINT(3113158514), "ETHERCAT_PLC1\_BASE\STRSOFTWAREVERSION",
1$UINT, TO_UDINT(3747917626), "WELCON_11\_BASE\_BASE\DEVICENAMESTR",
1$UINT, TO_UDINT(3734643842), "WELCON_11\_BASE\_BASE\PRODUCTREVSTR",
1$UINT, TO_UDINT(3719997469), "WELCON_21\_BASE\_BASE\DEVICENAMESTR",
1$UINT, TO_UDINT(3695453093), "WELCON_21\_BASE\_BASE\PRODUCTREVSTR",
1$UINT, TO_UDINT(3691992320), "WELCON_31\_BASE\_BASE\DEVICENAMESTR",
1$UINT, TO_UDINT(3723615928), "WELCON_31\_BASE\_BASE\PRODUCTREVSTR",
1$UINT, TO_UDINT(3624314451), "WELCON_41\_BASE\_BASE\DEVICENAMESTR",
1$UINT, TO_UDINT(3656920555), "WELCON_41\_BASE\_BASE\PRODUCTREVSTR",

_NO_ATTR, TO_UDINT(2395414379), "VARANMANAGER_11",

_NO_ATTR, TO_UDINT(3391823300), "WELCON_11",

_NO_ATTR, TO_UDINT(3775286791), "WELCON_21",

_NO_ATTR, TO_UDINT(4162682694), "WELCON_31",

_NO_ATTR, TO_UDINT(3076319617), "WELCON_41",

//Internal connections
0$UDINT,
45$UDINT,
TO_UDINT(5), "GetCILInterfacePLL", TO_UDINT(17),
TO_UDINT(7), "_SerLib1", TO_UDINT(2),
TO_UDINT(7), "_SerLib2", TO_UDINT(3),
TO_UDINT(7), "_CanLib1", TO_UDINT(0),
TO_UDINT(7), "_CanLib2", TO_UDINT(1),
TO_UDINT(7), "_SerLib3", TO_UDINT(4),
TO_UDINT(15), "GetCILInterface_ECAT", TO_UDINT(16),
TO_UDINT(15), "strSoftwareVersion", TO_UDINT(40),
TO_UDINT(15), "_SyncMeasureECAT1", TO_UDINT(5),
TO_UDINT(15), "EtherCAT_Hub_Base1", TO_UDINT(10),
TO_UDINT(24), "SafetyManager", TO_UDINT(35),
TO_UDINT(24), "HWRtPostScan", TO_UDINT(25),
TO_UDINT(24), "HwcLogging", TO_UDINT(23),
TO_UDINT(35), "UdpSendData", TO_UDINT(9),
TO_UDINT(35), "UdpReceiveData", TO_UDINT(8),
TO_UDINT(35), "SafetyRoutingTables1", TO_UDINT(36),
TO_UDINT(39), "SdiasManager1", TO_UDINT(38),
TO_UDINT(39), "SdiasHubBase1", TO_UDINT(37),
TO_UDINT(40), "MerkerEx0", TO_UDINT(26),
TO_UDINT(41), "MerkerEx0", TO_UDINT(27),
TO_UDINT(42), "MerkerEx0", TO_UDINT(28),
TO_UDINT(43), "MerkerEx0", TO_UDINT(29),
TO_UDINT(44), "MerkerEx0", TO_UDINT(30),
TO_UDINT(45), "MerkerEx0", TO_UDINT(31),
TO_UDINT(46), "MerkerEx0", TO_UDINT(32),
TO_UDINT(47), "MerkerEx0", TO_UDINT(33),
TO_UDINT(48), "MerkerEx0", TO_UDINT(34),
TO_UDINT(49), "ASCII_BIN1", TO_UDINT(6),
TO_UDINT(49), "Hub_Base_Root0", TO_UDINT(22),
TO_UDINT(50), "GetCILInterface_ECAT", TO_UDINT(18),
TO_UDINT(50), "DeviceNameStr", TO_UDINT(41),
TO_UDINT(50), "ProductRevStr", TO_UDINT(42),
TO_UDINT(50), "EtherCAT_Hub_Base_1", TO_UDINT(11),
TO_UDINT(51), "GetCILInterface_ECAT", TO_UDINT(19),
TO_UDINT(51), "DeviceNameStr", TO_UDINT(43),
TO_UDINT(51), "ProductRevStr", TO_UDINT(44),
TO_UDINT(51), "EtherCAT_Hub_Base_1", TO_UDINT(12),
TO_UDINT(52), "GetCILInterface_ECAT", TO_UDINT(20),
TO_UDINT(52), "DeviceNameStr", TO_UDINT(45),
TO_UDINT(52), "ProductRevStr", TO_UDINT(46),
TO_UDINT(52), "EtherCAT_Hub_Base_1", TO_UDINT(13),
TO_UDINT(53), "GetCILInterface_ECAT", TO_UDINT(21),
TO_UDINT(53), "DeviceNameStr", TO_UDINT(47),
TO_UDINT(53), "ProductRevStr", TO_UDINT(48),
TO_UDINT(53), "EtherCAT_Hub_Base_1", TO_UDINT(14),
0$UDINT,
27$UDINT,
TO_UDINT(7), "To_HwControl", TO_UDINT(24), "Control",
TO_UDINT(10), "toNextEtherCAT", TO_UDINT(15), "ClassState",
TO_UDINT(11), "toNextEtherCAT", TO_UDINT(50), "ClassState",
TO_UDINT(12), "toNextEtherCAT", TO_UDINT(51), "ClassState",
TO_UDINT(13), "toNextEtherCAT", TO_UDINT(52), "ClassState",
TO_UDINT(14), "toNextEtherCAT", TO_UDINT(53), "ClassState",
TO_UDINT(15), "ToHwControl", TO_UDINT(24), "Control",
TO_UDINT(22), "VaranConnect", TO_UDINT(49), "Control",
TO_UDINT(25), "toHwControlBase", TO_UDINT(24), "Control",
TO_UDINT(35), "To_HwControl", TO_UDINT(24), "Control",
TO_UDINT(37), "ToNextSDIAS", TO_UDINT(38), "ClassState",
TO_UDINT(38), "ToBusInterface", TO_UDINT(39), "CallCommand",
TO_UDINT(39), "ToHwControl", TO_UDINT(24), "Control",
TO_UDINT(40), "DataBuffer", TO_UDINT(26), "m_udLength",
TO_UDINT(41), "DataBuffer", TO_UDINT(27), "m_udLength",
TO_UDINT(42), "DataBuffer", TO_UDINT(28), "m_udLength",
TO_UDINT(43), "DataBuffer", TO_UDINT(29), "m_udLength",
TO_UDINT(44), "DataBuffer", TO_UDINT(30), "m_udLength",
TO_UDINT(45), "DataBuffer", TO_UDINT(31), "m_udLength",
TO_UDINT(46), "DataBuffer", TO_UDINT(32), "m_udLength",
TO_UDINT(47), "DataBuffer", TO_UDINT(33), "m_udLength",
TO_UDINT(48), "DataBuffer", TO_UDINT(34), "m_udLength",
TO_UDINT(49), "To_HwControl", TO_UDINT(24), "Control",
TO_UDINT(50), "toMaster", TO_UDINT(10), "ClassSvr",
TO_UDINT(51), "toMaster", TO_UDINT(11), "ClassSvr",
TO_UDINT(52), "toMaster", TO_UDINT(12), "ClassSvr",
TO_UDINT(53), "toMaster", TO_UDINT(13), "ClassSvr",

//Initialization values
0$UDINT,
86$UDINT,
TO_UDINT(0), "CanBus", TO_UDINT(1),//|HW_Network._base\CP313_IOs1\_CanLib1.CanBus;
TO_UDINT(1), "CanBus", TO_UDINT(2),//|HW_Network._base\CP313_IOs1\_CanLib2.CanBus;
TO_UDINT(2), "Com", TO_UDINT(1),//|HW_Network._base\CP313_IOs1\_SerLib1.Com;
TO_UDINT(3), "Com", TO_UDINT(2),//|HW_Network._base\CP313_IOs1\_SerLib2.Com;
TO_UDINT(4), "Com", TO_UDINT(3),//|HW_Network._base\CP313_IOs1\_SerLib3.Com;
TO_UDINT(5), "divisor", TO_UDINT(4),//|HW_Network._base\EtherCAT_PLC1\_SyncMeasureECAT1.divisor;
TO_UDINT(5), "PhaseRegDamping", TO_UDINT(0),//|HW_Network._base\EtherCAT_PLC1\_SyncMeasureECAT1.PhaseRegDamping;
TO_UDINT(10), "SplitterPlace", TO_UDINT(0),//|HW_Network.EtherCAT_PLC1\EtherCAT_Hub_Base1.SplitterPlace;
TO_UDINT(10), "BusType", TO_UDINT(0),//|HW_Network.EtherCAT_PLC1\EtherCAT_Hub_Base1.BusType;
TO_UDINT(11), "SplitterPlace", TO_UDINT(0),//|HW_Network.WELCON_11\EtherCAT_Hub_Base_1.SplitterPlace;
TO_UDINT(11), "BusType", TO_UDINT(0),//|HW_Network.WELCON_11\EtherCAT_Hub_Base_1.BusType;
TO_UDINT(12), "SplitterPlace", TO_UDINT(0),//|HW_Network.WELCON_21\EtherCAT_Hub_Base_1.SplitterPlace;
TO_UDINT(12), "BusType", TO_UDINT(0),//|HW_Network.WELCON_21\EtherCAT_Hub_Base_1.BusType;
TO_UDINT(13), "SplitterPlace", TO_UDINT(0),//|HW_Network.WELCON_31\EtherCAT_Hub_Base_1.SplitterPlace;
TO_UDINT(13), "BusType", TO_UDINT(0),//|HW_Network.WELCON_31\EtherCAT_Hub_Base_1.BusType;
TO_UDINT(14), "SplitterPlace", TO_UDINT(0),//|HW_Network.WELCON_41\EtherCAT_Hub_Base_1.SplitterPlace;
TO_UDINT(14), "BusType", TO_UDINT(0),//|HW_Network.WELCON_41\EtherCAT_Hub_Base_1.BusType;
TO_UDINT(15), "IsoStartPoint", TO_UDINT(50),//|HW_Network.EtherCAT_PLC1.IsoStartPoint;
TO_UDINT(15), "CoreSelect", TO_UDINT(0),//|HW_Network.EtherCAT_PLC1.CoreSelect;
TO_UDINT(15), "MasterID", TO_UDINT(1),//|HW_Network.EtherCAT_PLC1.MasterID;
TO_UDINT(15), "StateTransitionBehaviour", TO_UDINT(2#110),//|HW_Network.EtherCAT_PLC1.StateTransitionBehaviour;
TO_UDINT(15), "StateTransitionTimeout", TO_UDINT(20000),//|HW_Network.EtherCAT_PLC1.StateTransitionTimeout;
TO_UDINT(15), "SynchronizationMode", TO_UDINT(0),//|HW_Network.EtherCAT_PLC1.SynchronizationMode;
TO_UDINT(15), "PhaseRegDamping", TO_UDINT(0),//|HW_Network.EtherCAT_PLC1.PhaseRegDamping;
TO_UDINT(15), "MissingFrameBehaviour", TO_UDINT(3),//|HW_Network.EtherCAT_PLC1.MissingFrameBehaviour;
TO_UDINT(22), "Splitter_Place", TO_UDINT(0),//|HW_Network.VaranManager_11\Hub_Base_Root0.Splitter_Place;
TO_UDINT(24), "UdpSafetyPort", TO_UDINT(10823),//|HW_Network.HwControl1.UdpSafetyPort;
TO_UDINT(24), "InterfaceNo", TO_UDINT(1),//|HW_Network.HwControl1.InterfaceNo;
TO_UDINT(24), "RtTaskSync", TO_UDINT(0),//|HW_Network.HwControl1.RtTaskSync;
TO_UDINT(26), "ThreadSafe", TO_UDINT(0),//|HW_Network.strSoftwareVersion\_base\EtherCAT_PLC1\MerkerEx0.ThreadSafe;
TO_UDINT(27), "ThreadSafe", TO_UDINT(0),//|HW_Network.DeviceNameStr\_base\_base\WELCON_11\MerkerEx0.ThreadSafe;
TO_UDINT(28), "ThreadSafe", TO_UDINT(0),//|HW_Network.ProductRevStr\_base\_base\WELCON_11\MerkerEx0.ThreadSafe;
TO_UDINT(29), "ThreadSafe", TO_UDINT(0),//|HW_Network.DeviceNameStr\_base\_base\WELCON_21\MerkerEx0.ThreadSafe;
TO_UDINT(30), "ThreadSafe", TO_UDINT(0),//|HW_Network.ProductRevStr\_base\_base\WELCON_21\MerkerEx0.ThreadSafe;
TO_UDINT(31), "ThreadSafe", TO_UDINT(0),//|HW_Network.DeviceNameStr\_base\_base\WELCON_31\MerkerEx0.ThreadSafe;
TO_UDINT(32), "ThreadSafe", TO_UDINT(0),//|HW_Network.ProductRevStr\_base\_base\WELCON_31\MerkerEx0.ThreadSafe;
TO_UDINT(33), "ThreadSafe", TO_UDINT(0),//|HW_Network.DeviceNameStr\_base\_base\WELCON_41\MerkerEx0.ThreadSafe;
TO_UDINT(34), "ThreadSafe", TO_UDINT(0),//|HW_Network.ProductRevStr\_base\_base\WELCON_41\MerkerEx0.ThreadSafe;
TO_UDINT(35), "UdpSafetyPort", TO_UDINT(10823),//|HW_Network.HwControl1\SafetyManager.UdpSafetyPort;
TO_UDINT(35), "InterfaceNo", TO_UDINT(1),//|HW_Network.HwControl1\SafetyManager.InterfaceNo;
TO_UDINT(35), "UdpSafetyRequestCycle", TO_UDINT(UDP_MIN_REQUEST_TIME),//|HW_Network.HwControl1\SafetyManager.UdpSafetyRequestCycle;
TO_UDINT(35), "UdpSafetyResponseTimeout", TO_UDINT(UDP_MIN_RESPONSE_TIMEOUT),//|HW_Network.HwControl1\SafetyManager.UdpSafetyResponseTimeout;
TO_UDINT(37), "SplitterPlace", TO_UDINT(0),//|HW_Network.SdiasPLC1\SdiasHubBase1.SplitterPlace;
TO_UDINT(38), "DeviceID", TO_UDINT(0),//|HW_Network.SdiasPLC1\SdiasManager1.DeviceID;
TO_UDINT(38), "AutoFarMem", TO_UDINT(0),//|HW_Network.SdiasPLC1\SdiasManager1.AutoFarMem;
TO_UDINT(39), "CycleTime", TO_UDINT(1000),//|HW_Network.SdiasPLC1.CycleTime;
TO_UDINT(39), "IsoStartPoint", TO_UDINT(50),//|HW_Network.SdiasPLC1.IsoStartPoint;
TO_UDINT(39), "AutoFarMem", TO_UDINT(0),//|HW_Network.SdiasPLC1.AutoFarMem;
TO_UDINT(40), "SingleRealloc", TO_UDINT(1),//|HW_Network._base\EtherCAT_PLC1\strSoftwareVersion.SingleRealloc;
TO_UDINT(41), "SingleRealloc", TO_UDINT(1),//|HW_Network._base\_base\WELCON_11\DeviceNameStr.SingleRealloc;
TO_UDINT(42), "SingleRealloc", TO_UDINT(1),//|HW_Network._base\_base\WELCON_11\ProductRevStr.SingleRealloc;
TO_UDINT(43), "SingleRealloc", TO_UDINT(1),//|HW_Network._base\_base\WELCON_21\DeviceNameStr.SingleRealloc;
TO_UDINT(44), "SingleRealloc", TO_UDINT(1),//|HW_Network._base\_base\WELCON_21\ProductRevStr.SingleRealloc;
TO_UDINT(45), "SingleRealloc", TO_UDINT(1),//|HW_Network._base\_base\WELCON_31\DeviceNameStr.SingleRealloc;
TO_UDINT(46), "SingleRealloc", TO_UDINT(1),//|HW_Network._base\_base\WELCON_31\ProductRevStr.SingleRealloc;
TO_UDINT(47), "SingleRealloc", TO_UDINT(1),//|HW_Network._base\_base\WELCON_41\DeviceNameStr.SingleRealloc;
TO_UDINT(48), "SingleRealloc", TO_UDINT(1),//|HW_Network._base\_base\WELCON_41\ProductRevStr.SingleRealloc;
TO_UDINT(49), "VaranManagerTime", TO_UDINT(1000000),//|HW_Network.VaranManager_11.VaranManagerTime;
TO_UDINT(49), "VaranManagerNr", TO_UDINT(0),//|HW_Network.VaranManager_11.VaranManagerNr;
TO_UDINT(49), "PayloadFrame", TO_UDINT(0),//|HW_Network.VaranManager_11.PayloadFrame;
TO_UDINT(49), "CoreSelect", TO_UDINT(0),//|HW_Network.VaranManager_11.CoreSelect;
TO_UDINT(49), "InterframeGap", TO_UDINT(0),//|HW_Network.VaranManager_11.InterframeGap;
TO_UDINT(50), "SlaveIndex", TO_UDINT(0),//|HW_Network.WELCON_11.SlaveIndex;
TO_UDINT(50), "Required", TO_UDINT(1),//|HW_Network.WELCON_11.Required;
TO_UDINT(50), "NoSDOBuffer", TO_UDINT(0),//|HW_Network.WELCON_11.NoSDOBuffer;
TO_UDINT(50), "NoAsyncBuffer", TO_UDINT(0),//|HW_Network.WELCON_11.NoAsyncBuffer;
TO_UDINT(50), "NoSSCBuffer", TO_UDINT(0),//|HW_Network.WELCON_11.NoSSCBuffer;
TO_UDINT(50), "UseDefaultEnableSequence", TO_UDINT(1),//|HW_Network.WELCON_11.UseDefaultEnableSequence;
TO_UDINT(51), "SlaveIndex", TO_UDINT(1),//|HW_Network.WELCON_21.SlaveIndex;
TO_UDINT(51), "Required", TO_UDINT(1),//|HW_Network.WELCON_21.Required;
TO_UDINT(51), "NoSDOBuffer", TO_UDINT(0),//|HW_Network.WELCON_21.NoSDOBuffer;
TO_UDINT(51), "NoAsyncBuffer", TO_UDINT(0),//|HW_Network.WELCON_21.NoAsyncBuffer;
TO_UDINT(51), "NoSSCBuffer", TO_UDINT(0),//|HW_Network.WELCON_21.NoSSCBuffer;
TO_UDINT(51), "UseDefaultEnableSequence", TO_UDINT(1),//|HW_Network.WELCON_21.UseDefaultEnableSequence;
TO_UDINT(52), "SlaveIndex", TO_UDINT(2),//|HW_Network.WELCON_31.SlaveIndex;
TO_UDINT(52), "Required", TO_UDINT(1),//|HW_Network.WELCON_31.Required;
TO_UDINT(52), "NoSDOBuffer", TO_UDINT(0),//|HW_Network.WELCON_31.NoSDOBuffer;
TO_UDINT(52), "NoAsyncBuffer", TO_UDINT(0),//|HW_Network.WELCON_31.NoAsyncBuffer;
TO_UDINT(52), "NoSSCBuffer", TO_UDINT(0),//|HW_Network.WELCON_31.NoSSCBuffer;
TO_UDINT(52), "UseDefaultEnableSequence", TO_UDINT(1),//|HW_Network.WELCON_31.UseDefaultEnableSequence;
TO_UDINT(53), "SlaveIndex", TO_UDINT(3),//|HW_Network.WELCON_41.SlaveIndex;
TO_UDINT(53), "Required", TO_UDINT(1),//|HW_Network.WELCON_41.Required;
TO_UDINT(53), "NoSDOBuffer", TO_UDINT(0),//|HW_Network.WELCON_41.NoSDOBuffer;
TO_UDINT(53), "NoAsyncBuffer", TO_UDINT(0),//|HW_Network.WELCON_41.NoAsyncBuffer;
TO_UDINT(53), "NoSSCBuffer", TO_UDINT(0),//|HW_Network.WELCON_41.NoSSCBuffer;
TO_UDINT(53), "UseDefaultEnableSequence", TO_UDINT(1),//|HW_Network.WELCON_41.UseDefaultEnableSequence;

//Symbolic initialization values
0$UDINT,
0$UDINT,

//Initialization of string values
0$UDINT,
0$UDINT,

//Configuration of tasks (RealTime, Cyclic, Background)
0$UDINT,
1$UDINT,
TO_UDINT(25), (1)$UDINT, 4194304$DINT, 	//HWCONTROL1\HWRTPOSTSCAN

0$UDINT,
0$UDINT,

0$UDINT,
0$UDINT,

//External connections
0$UDINT,
0$UDINT,

//Magic internal connections
0$UDINT,
5$UDINT,
TO_UDINT(5), "PhaseRegDamping", TO_UDINT(15), "PhaseRegDamping",
TO_UDINT(35), "UdpSafetyPort", TO_UDINT(24), "UdpSafetyPort",
TO_UDINT(35), "InterfaceNo", TO_UDINT(24), "InterfaceNo",
TO_UDINT(35), "SafetyDomainTimeout", TO_UDINT(24), "SafetyDomainTimeout",
TO_UDINT(38), "AutoFarMem", TO_UDINT(39), "AutoFarMem",

//Configuration of timeslots of tasks (RealTime, Cyclic)
#ifdef __LSLLDR_TIMESLOTS__
0$UDINT,
0$UDINT,

0$UDINT,
0$UDINT,

#endif //__LSLLDR_TIMESLOTS__

//MultiMaster connections
#ifdef __LSLLDR_MULTIMASTER__
0$UDINT,
0$UDINT,
#endif //__LSLLDR_MULTIMASTER__

//Configuration for task ID (RealTime, CyclicTime)
#ifdef __LSLLDR_TASKID__
"\\\\TASKS2  "
0$UDINT,
1$UDINT,
(0)$UDINT, 	//HWCONTROL1\HWRTPOSTSCAN

0$UDINT,
0$UDINT,

0$UDINT,
0$UDINT,

#endif //__LSLLDR_TASKID__

END_FUNCTION
